Fanuc KAREL source: KO00098.KL

PROGRAM KO00098
%NOLOCKGROUP
VAR
  A: INTEGER
  B: INTEGER
  OUT: REAL
BEGIN
  A = 1
  B = 2
  OUT = ATAN2(A, B)
END KO00098
